TYPE ST_ValveStatus :
STRUCT
	eState		: E_ValveState;
	bInterlocked	: BOOL;
	nCycles		: UDINT;
	fOpenTime	: LREAL; // s
END_STRUCT
END_TYPE

(* stored: Version 1.1.0.1
   DUT ST_ValveStatus: Id {a826fa27-fbb9-47d0-9d7e-3596e5163cef} *)
